FUNCTION F_Total : UDINT
VAR_IN_OUT
    counts : ARRAY[*] OF UDINT;
END_VAR
VAR
    i : DINT;
END_VAR


F_Total := 0;
FOR i := LOWER_BOUND(counts, 1) TO UPPER_BOUND(counts, 1) DO
    F_Total := F_Total + counts[i];
END_FOR;

END_FUNCTION

(* stored: Version 1.1.0.1, ProductVersion 3.1 *)
